(* IEC 61131-3 sources: auto-inspection-station/plc/openplc_project/pous/programs, 1 file *)

(* ---- status_logic.st ---- *)
PROGRAM status_logic
  VAR
    SIM_MODE : BOOL;
  END_VAR

// IF SIM_MODE THEN
//     IN_UNIT_SERIAL := SIM_UNIT_SERIAL_IN;
//     IN_FAIL_REASON := SIM_FAIL_REASON_IN;
// ELSE
//     IN_UNIT_SERIAL := 0;
//     IN_FAIL_REASON := 0;
// END_IF;

// IF S_IDLE THEN
//     STATE_CODE := 0;
// ELSIF S_READY THEN
//     STATE_CODE := 10;
// ELSIF S_INSPECTING THEN
//     STATE_CODE := 20;
// ELSIF S_PASS_RELEASE THEN
//     STATE_CODE := 30;
// ELSIF S_REJECT_EXTEND THEN
//     STATE_CODE := 40;
// ELSIF S_REJECT_RETRACT THEN
//     STATE_CODE := 50;
// ELSIF S_FAULT THEN
//     STATE_CODE := 90;
// END_IF;

// IF UNIT_RISE THEN
//     CURRENT_SERIAL := IN_UNIT_SERIAL;
//     CYCLE_START_MS := SCENARIO_STEP;
// END_IF;

// IF RESULT_FAIL_LATCH AND NOT RESULT_PASS_LATCH THEN
//     CURRENT_FAIL_REASON := IN_FAIL_REASON;
// ELSIF RESULT_PASS_LATCH THEN
//     CURRENT_FAIL_REASON := 0;
// END_IF;

// IF PASS_COMPLETE_PULSE THEN
//     TOTAL_UNITS := TOTAL_UNITS + 1;
//     LAST_SERIAL := CURRENT_SERIAL;
//     LAST_RESULT := 1;
//     LAST_FAIL_REASON := 0;
//     LAST_CYCLE_TIME_MS := SCENARIO_STEP - CYCLE_START_MS;
// END_IF;

// IF FAIL_COMPLETE_PULSE THEN
//     TOTAL_UNITS := TOTAL_UNITS + 1;
//     TOTAL_REJECTS := TOTAL_REJECTS + 1;
//     LAST_SERIAL := CURRENT_SERIAL;
//     LAST_RESULT := 2;
//     LAST_FAIL_REASON := CURRENT_FAIL_REASON;
//     LAST_CYCLE_TIME_MS := SCENARIO_STEP - CYCLE_START_MS;
// END_IF;

// IF FAULT_ESTOP THEN
//     FAULT_CODE := 100;
// ELSIF FAULT_GUARD THEN
//     FAULT_CODE := 110;
// ELSIF FAULT_EXTEND_TIMEOUT THEN
//     FAULT_CODE := 120;
// ELSIF FAULT_RETRACT_TIMEOUT THEN
//     FAULT_CODE := 130;
// ELSIF FAULT_UNIT_STUCK THEN
//     FAULT_CODE := 140;
// ELSIF FAULT_VISION_UNSTABLE THEN
//     FAULT_CODE := 150;
// ELSIF FAULT_OUTPUT_CONFLICT THEN
//     FAULT_CODE := 160;
// ELSE
//     FAULT_CODE := 0;
// END_IF;

END_PROGRAM
